(* PLC project , Example Fixture *)

PROGRAM Check
  VAR_INPUT
    Level : REAL;
  END_VAR
  VAR_OUTPUT
    Full : BOOL;
  END_VAR

(* FBD diagram, written out as Structured Text *)
Full := Level = 2.5;
END_PROGRAM

CONFIGURATION c
  RESOURCE r ON PLC
  END_RESOURCE
END_CONFIGURATION
